Fanuc KAREL source: KT00903.KL

PROGRAM KT00903
%NOLOCKGROUP
%ENVIRONMENT VECTR
VAR
  P1: POSITION
  P2: POSITION
  OUT: VECTOR
BEGIN
  OUT = APPROACH(P1)
END KT00903
